(* IEC 61131-3 sources: plcfuzz/testcases/beremiz_projects/blank_code, 1 file *)

(* ---- blank.st ---- *)
PROGRAM program0
  VAR
    LED AT %QX0.0 : BOOL;
  END_VAR

  LED := TRUE;
END_PROGRAM

CONFIGURATION Config0

  RESOURCE Res0 ON PLC
    TASK task0(INTERVAL := T#20ms,PRIORITY := 0);
    PROGRAM instance0 WITH task0 : program0;
  END_RESOURCE
END_CONFIGURATION
